FUNCTION_BLOCK normalise1 (* Basic Function Block Type *)
  (* Standard: 61499-2 *)
  (* Version 0.0, 12/26/2019, prana, nxtControl GmbH, Template *)
  PACKAGE Main;
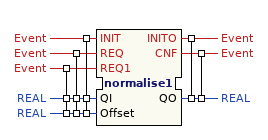
  EVENT_INPUT
    INIT WITH QI, Offset; (* Initialization Request *)
    REQ WITH QI, Offset; (* Normal Execution Request *)
    REQ1 WITH QI, Offset;
  END_EVENT
  EVENT_OUTPUT
    INITO WITH QO; (* Initialization Confirm *)
    CNF WITH QO; (* Execution Confirmation *)
  END_EVENT
  VAR_INPUT
    QI : REAL; (* Input event qualifier *)
    Offset : REAL;
  END_VAR
  VAR_OUTPUT
    QO : REAL; (* Output event qualifier *)
  END_VAR
  VAR
    QI1 : REAL;
  END_VAR
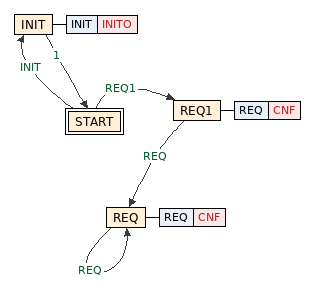
  EC_STATES
    START; (* Initial State *)
    REQ : REQ -> CNF; (* Normal execution *)
    REQ1 : REQ -> CNF;
    INIT : INIT -> INITO;
  END_STATES
  EC_TRANSITIONS
    REQ1 TO REQ := REQ;
    REQ TO REQ := REQ;
    START TO REQ1 := REQ1;
    INIT TO START := 1;
    START TO INIT := INIT;
  END_TRANSITIONS
  ALGORITHM INIT IN ST: (* Initialization algorithm *)
;
  END_ALGORITHM
  ALGORITHM REQ IN ST: (* Normally executed algorithm *)
QI1 := QI - Offset;
QO := ( QI1 - 120 ) / ( 260) ;
  END_ALGORITHM
END_FUNCTION_BLOCK
